Fanuc KAREL source: KA00036.KL

PROGRAM KA00036
%NOLOCKGROUP
VAR
  SRC: BOOLEAN
  DST: ARRAY[2] OF SHORT
BEGIN
  SRC = TRUE
  DST[1] = SRC
END KA00036
